(* IEC 61131-3 sources: tinyplc/examples, 3 files *)

(* ---- button_led.st ---- *)
PROGRAM Main
VAR_INPUT
    BTN : BOOL;
END_VAR
VAR_OUTPUT
    LED : BOOL;
END_VAR
VAR
    n : DINT;
END_VAR
(* n increments every scan while BTN is TRUE, not once per press. *)
IF BTN THEN
    n := n + 1;
END_IF;
LED := NOT BTN;
END_PROGRAM

(* ---- download_led_off.st ---- *)
(* Serial-download demonstration. Tags deliberately differ from boot ordering.
   When BTN is released LD2 is OFF; activation starts N from zero. *)
PROGRAM Downloaded
VAR N : DINT; END_VAR
VAR_INPUT BTN : BOOL; END_VAR
VAR_OUTPUT LED : BOOL; END_VAR
N := N + 1;
LED := BTN;
END_PROGRAM

(* ---- ton_led.st ---- *)
PROGRAM DelayedButton
VAR_INPUT BTN : BOOL; END_VAR
VAR_OUTPUT LED : BOOL; END_VAR
VAR Delay : TON; END_VAR
Delay(IN := BTN, PT := T#500ms);
LED := Delay.Q;
END_PROGRAM
